RoboDK station: TMflow export test.rdk

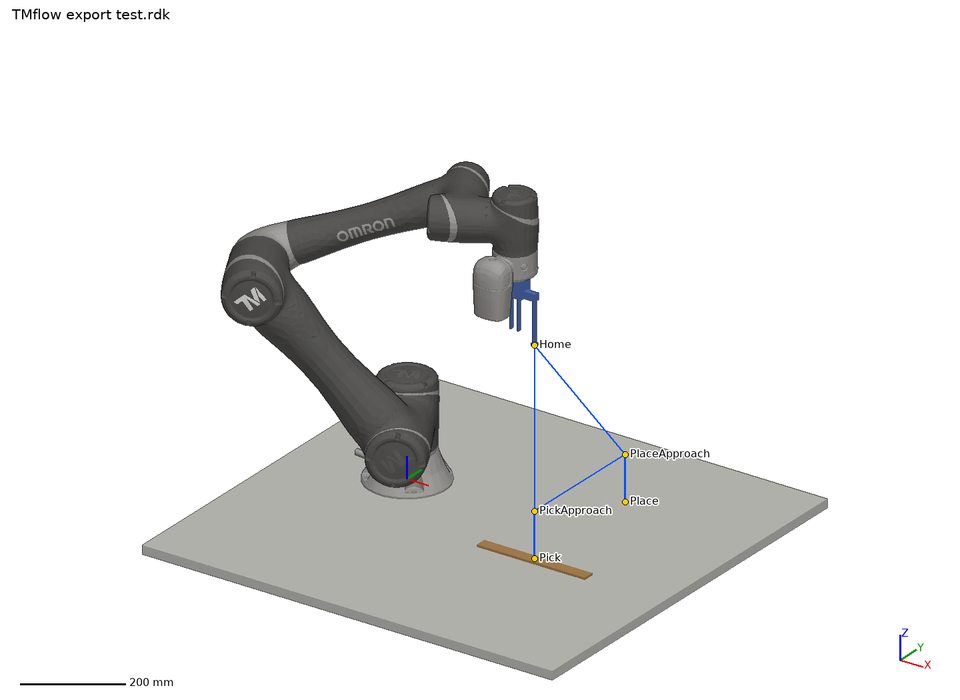
[picture v0: the station drawn from its stored meshes, robots at their saved joint values, targets as dots, program paths as lines]
Station TMflow export test (saved by RoboDK 6.1.1). Poses are relative to the parent item; angles as X-Y-Z fixed-axis rotations.
  - frame Cell at (0, 0, 0) mm
    - object Table at (0, 0, 0) mm, size 950 x 910 x 19 mm
    - frame Omron TM5-900 Base at (0, 0, 0) mm
      - robot Omron TM5-900: 6 axes, payload 4 kg, reach 900 mm, repeatability 0.05 mm, weight 22.6 kg
          modified DH rows (alpha deg, a mm, theta deg, d mm): 0, 0, 0, 145.2; 90, 0, 90, 0; 0, 429, 0, 0; 0, 411, -90, 122.3; -90, 0, 0, 106.5; 90, 0, 180, 114.15
          joint limits [-270, -180, -155, -180, -180, -270] to [270, 180, 155, 180, 180, 270]; home [0, 0, 90, -90, 90, 0]; saved at [29.3, -39.9, 110, 19.9, 90, 119.3]
        - tool Vacuum, TCP at (45, 0, 135) mm, size 75 x 30 x 135 mm
    - object Plank at (400, -150, -1) mm, rotated rx 0 ry 0 rz 90 deg, size 25 x 250 x 5 mm, geometry from plank.stl
    - target Home (joint target) at (294.77, -0.08, 365.06) mm, rotated rx -180 ry 0 rz 0 deg; joints [29.3, -39.9, 110, 19.9, 90, 119.3] of Omron TM5-900
    - target PickApproach (Cartesian target) at (400, -150, 104) mm, rotated rx 180 ry 0 rz 0 deg; joints [-4.404, -12.65, 133.481, -30.83, 90, 85.596] of Omron TM5-900
    - target Pick (Cartesian target) at (400, -150, 4) mm, rotated rx 180 ry 0 rz 0 deg; joints [-4.404, 0.314, 141.05, -51.364, 90, 85.596] of Omron TM5-900
    - target PlaceApproach (Cartesian target) at (400, 150, 104) mm, rotated rx 180 ry 0 rz 0 deg; joints [41.408, -12.65, 133.481, -30.83, 90, 131.408] of Omron TM5-900
    - target Place (Cartesian target) at (400, 150, 4) mm, rotated rx 180 ry 0 rz 0 deg; joints [41.408, 0.314, 141.05, -51.364, 90, 131.408] of Omron TM5-900
  - program PickPlaceTest (19 instructions, listed below)
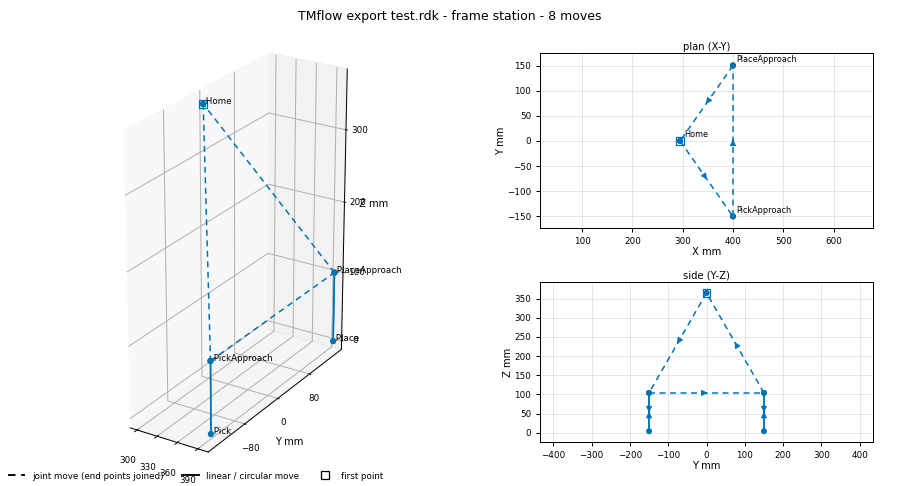
[picture p0: tool path of TMflow export test.rdk in frame station, 8 of 8 moves have a stored position in this frame; points joined in program order, loops and branches not executed]

--- program PickPlaceTest (robot Omron TM5-900) ---
  Simulation: plank to start
  Set Ref.: Cell
  Set Tool: Vacuum
  Set speed (100.0 mm/s)
  Smooth(0)
  MoveJ (Home)
  MoveJ (PickApproach)
  MoveL (Pick)
  Set IO_0=1
  Simulation: attach plank
  Pause 500 ms
  MoveL (PickApproach)
  MoveJ (PlaceApproach)
  MoveL (Place)
  Set IO_0=0
  Simulation: release plank
  Pause 500 ms
  MoveL (PlaceApproach)
  MoveJ (Home)
